{attribute 'no_assign'}
FUNCTION_BLOCK FB_LN_WTURBINE_LD0_WPPD1 EXTENDS FB_AcsiCommonLogicalNodeClass
VAR_INPUT
	Beh: FB_DO_WTURBINE_LD0_WPPD1_Beh := (sClass:='ENS', bLinkResult:=THIS^.AddDataToContainer(ipData:=Beh));
	DevSt: FB_DO_WTURBINE_LD0_WPPD1_DevSt := (sClass:='STV', bLinkResult:=THIS^.AddDataToContainer(ipData:=DevSt));
	DevOp: FB_DO_WTURBINE_LD0_WPPD1_DevOp := (sClass:='CMD', bLinkResult:=THIS^.AddDataToContainer(ipData:=DevOp));
	ClrOp: FB_DO_WTURBINE_LD0_WPPD1_ClrOp := (sClass:='CMD', bLinkResult:=THIS^.AddDataToContainer(ipData:=ClrOp));
	
	ds01: FB_DS_TEMPLATE_LD1_WPPD1_ds01 := (bLinkResult:=THIS^.AddDataSetToContainer(ipDataSet:=ds01));
	
	urcb01: FB_ScsmUrCBImplClass := (RptID:=(sValue:='WTURBINELD0/WPPD1.urcb01'), DatSet:=(sValue:='WTURBINELD0/WPPD1.ds01'), OptFlds:=(SequenceNumber:=FALSE, ReportTimeStamp:=FALSE, ReasonForInclusion:=FALSE, DataSetName:=FALSE, DataReference:=FALSE, BufferOverflow:=FALSE, EntryID:=FALSE, ConfRevision:=FALSE), TrgOps:=(DataChange:=FALSE, QualityChange:=FALSE, DataUpdate:=FALSE, Integrity:=FALSE, GeneralInterrogation:=TRUE), bLinkResult:=THIS^.AddUnbufferedReportControlBlockToContainer(ipUnbufferedReportControlBlock:=urcb01));
END_VAR
VAR
END_VAR

END_FUNCTION_BLOCK

(* stored: Version 1.1.0.1
   POU FB_LN_WTURBINE_LD0_WPPD1: Id {1c0b0c0f-c62d-4c7c-afae-67772457a8f7}, SpecialFunc None *)
